FUNCTION_BLOCK AOption_EVENT_TO_X (* Composite FB for convert EVENT to AOption (Fan-Out, haelt den PLUG) *)
  (* Standard: 61499-2; Description: Copyright (c) 2026 Meisterschulen am Ostbahnhof This program and the accompanying materials are made available under the terms of the Eclipse Public License 2.0 which is available at https://www.eclipse.org/legal/epl-2.0/ SPDX-License-Identifier: EPL-2.0 *)
  (* Version 1.0, 2026-10-13, Franz Höpfinger, Meisterschulen am Ostbahnhof *)
  PACKAGE Option::conversion;
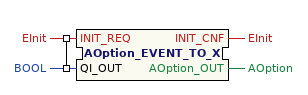
  EVENT_INPUT
    INIT_REQ : EInit WITH QI_OUT; (* Request to Adapter *)
  END_EVENT
  EVENT_OUTPUT
    INIT_CNF : EInit; (* Confirmation from Adapter *)
  END_EVENT
  VAR_INPUT
    QI_OUT : BOOL; (* Event Input Qualifier (IEC 61499-1): TRUE=Option anfordern/aktivieren, FALSE=zurueckziehen *)
  END_VAR
  PLUGS
    AOption_OUT : Option::AOption; (* Adapter Output *)
  END_PLUGS
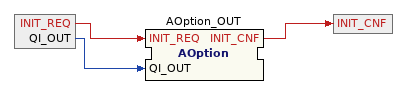
  EVENT_CONNECTIONS
    INIT_REQ TO AOption_OUT.INIT_REQ;
    AOption_OUT.INIT_CNF TO INIT_CNF;
  END_CONNECTIONS
  DATA_CONNECTIONS
    QI_OUT TO AOption_OUT.QI_OUT;
  END_CONNECTIONS
END_FUNCTION_BLOCK
